(* IEC 61131-3 sources: Industrial-automation-using-LLMs/datasets/Industrial_data/test_harness/test_case (part 2) *)

(* ---- SEQUENCE_8_TestCases (1).st ---- *)
FUNCTION_BLOCK FB_TEST_0
  VAR_OUTPUT
    Finished : BOOL;
    Failed : BOOL;
  END_VAR
  VAR
    TestBlock : SEQUENCE_8;
    TestState : INT;
    Timer : TON;
  END_VAR

  Timer(IN:=TRUE, PT:= T#0s); (* placeholder for later usage *)

  CASE testState OF
    0:
      IF (Timer.Q) THEN
        TestBlock(IN0 := TRUE, IN1 := TRUE, IN2 := TRUE, IN3 := TRUE, IN4 := TRUE, IN5 := TRUE, IN6 := TRUE, IN7 := TRUE, START := FALSE, RST := TRUE, STOP_ON_ERROR := TRUE);
        TestState:=TestState+1;
      END_IF;
      Timer(IN:=TRUE, PT:=T#0s);
    1:
      IF (Timer.Q) THEN
      {printf("0,0: TestBlock.Q0 = FALSE  actual=%lf\n", (double)__GET_VAR(data__->TESTBLOCK.Q0,));}
      {printf("0,0: TestBlock.Q1 = FALSE  actual=%lf\n", (double)__GET_VAR(data__->TESTBLOCK.Q1,));}
      {printf("0,0: TestBlock.Q2 = FALSE  actual=%lf\n", (double)__GET_VAR(data__->TESTBLOCK.Q2,));}
      {printf("0,0: TestBlock.Q3 = FALSE  actual=%lf\n", (double)__GET_VAR(data__->TESTBLOCK.Q3,));}
      {printf("0,0: TestBlock.Q4 = FALSE  actual=%lf\n", (double)__GET_VAR(data__->TESTBLOCK.Q4,));}
      {printf("0,0: TestBlock.Q5 = FALSE  actual=%lf\n", (double)__GET_VAR(data__->TESTBLOCK.Q5,));}
      {printf("0,0: TestBlock.Q6 = FALSE  actual=%lf\n", (double)__GET_VAR(data__->TESTBLOCK.Q6,));}
      {printf("0,0: TestBlock.Q7 = FALSE  actual=%lf\n", (double)__GET_VAR(data__->TESTBLOCK.Q7,));}
      {printf("0,0: TestBlock.QX = FALSE  actual=%lf\n", (double)__GET_VAR(data__->TESTBLOCK.QX,));}
      {printf("0,0: TestBlock.RUN = FALSE  actual=%lf\n", (double)__GET_VAR(data__->TESTBLOCK.RUN,));}
      {printf("0,0: TestBlock._STEP = -1  actual=%lf\n", (double)__GET_VAR(data__->TESTBLOCK._STEP,));}
      {printf("0,0: TestBlock.STATUS = 110  actual=%lf\n", (double)__GET_VAR(data__->TESTBLOCK.STATUS,));}
        IF NOT(TestBlock.Q0 = FALSE AND TestBlock.Q1 = FALSE AND TestBlock.Q2 = FALSE AND TestBlock.Q3 = FALSE AND TestBlock.Q4 = FALSE AND TestBlock.Q5 = FALSE AND TestBlock.Q6 = FALSE AND TestBlock.Q7 = FALSE AND TestBlock.QX = FALSE AND TestBlock.RUN = FALSE AND TestBlock._STEP = -1 AND TestBlock.STATUS = 110) THEN Failed := TRUE; END_IF;
      END_IF;
      Finished:=TRUE;
  END_CASE;
END_FUNCTION_BLOCK

FUNCTION_BLOCK FB_TEST_1
  VAR_OUTPUT
    Finished : BOOL;
    Failed : BOOL;
  END_VAR
  VAR
    TestBlock : SEQUENCE_8;
    TestState : INT;
    Timer : TON;
  END_VAR

  Timer(IN:=TRUE, PT:= T#0s); (* placeholder for later usage *)

  CASE testState OF
    0:
      IF (Timer.Q) THEN
        TestBlock(IN0 := TRUE, IN1 := TRUE, IN2 := TRUE, IN3 := TRUE, IN4 := TRUE, IN5 := TRUE, IN6 := TRUE, IN7 := TRUE, START := TRUE, RST := FALSE, STOP_ON_ERROR := FALSE);
        TestState:=TestState+1;
      END_IF;
      Timer(IN:=TRUE, PT:=T#0s);
    1:
      IF (Timer.Q) THEN
      {printf("1,0: TestBlock.Q0 = TRUE  actual=%lf\n", (double)__GET_VAR(data__->TESTBLOCK.Q0,));}
      {printf("1,0: TestBlock.Q1 = FALSE  actual=%lf\n", (double)__GET_VAR(data__->TESTBLOCK.Q1,));}
      {printf("1,0: TestBlock.Q2 = FALSE  actual=%lf\n", (double)__GET_VAR(data__->TESTBLOCK.Q2,));}
      {printf("1,0: TestBlock.Q3 = FALSE  actual=%lf\n", (double)__GET_VAR(data__->TESTBLOCK.Q3,));}
      {printf("1,0: TestBlock.Q4 = FALSE  actual=%lf\n", (double)__GET_VAR(data__->TESTBLOCK.Q4,));}
      {printf("1,0: TestBlock.Q5 = FALSE  actual=%lf\n", (double)__GET_VAR(data__->TESTBLOCK.Q5,));}
      {printf("1,0: TestBlock.Q6 = FALSE  actual=%lf\n", (double)__GET_VAR(data__->TESTBLOCK.Q6,));}
      {printf("1,0: TestBlock.Q7 = FALSE  actual=%lf\n", (double)__GET_VAR(data__->TESTBLOCK.Q7,));}
      {printf("1,0: TestBlock.QX = TRUE  actual=%lf\n", (double)__GET_VAR(data__->TESTBLOCK.QX,));}
      {printf("1,0: TestBlock.RUN = TRUE  actual=%lf\n", (double)__GET_VAR(data__->TESTBLOCK.RUN,));}
      {printf("1,0: TestBlock._STEP = 0  actual=%lf\n", (double)__GET_VAR(data__->TESTBLOCK._STEP,));}
      {printf("1,0: TestBlock.STATUS = 111  actual=%lf\n", (double)__GET_VAR(data__->TESTBLOCK.STATUS,));}
        IF NOT(TestBlock.Q0 = TRUE AND TestBlock.Q1 = FALSE AND TestBlock.Q2 = FALSE AND TestBlock.Q3 = FALSE AND TestBlock.Q4 = FALSE AND TestBlock.Q5 = FALSE AND TestBlock.Q6 = FALSE AND TestBlock.Q7 = FALSE AND TestBlock.QX = TRUE AND TestBlock.RUN = TRUE AND TestBlock._STEP = 0 AND TestBlock.STATUS = 111) THEN Failed := TRUE; END_IF;
      END_IF;
      Finished:=TRUE;
  END_CASE;
END_FUNCTION_BLOCK

PROGRAM TestRunnerProgram
VAR
  testResult AT %QX0.0 : BOOL := FALSE;
END_VAR
VAR
  totalTests AT %QW0 : INT := 0;
  passedTests AT %QW1 : INT := 0;
END_VAR
VAR
  i: INT := 0;
  testOutcomeArray : ARRAY [0..1] OF BOOL;
  Test_0: FB_TEST_0;
  Test_1: FB_TEST_1;
END_VAR

  IF NOT Test_0.Finished AND NOT Test_0.FAILED THEN totalTests := totalTests + 1; Test_0(); END_IF;
  IF Test_0.Finished THEN testOutcomeArray[0] := TRUE; END_IF;
  IF NOT Test_1.Finished AND NOT Test_1.FAILED THEN totalTests := totalTests + 1; Test_1(); END_IF;
  IF Test_1.Finished THEN testOutcomeArray[1] := TRUE; END_IF;

  passedTests := 0;
  FOR i:=0 TO 1 DO
    IF testOutcomeArray[i]=TRUE THEN passedTests := passedTests+1; END_IF;
  END_FOR;
END_PROGRAM

(* ---- SEQUENCE_8_TestCases.st ---- *)
FUNCTION_BLOCK FB_TEST_0
  VAR_OUTPUT
    Finished : BOOL;
    Failed : BOOL;
  END_VAR
  VAR
    TestBlock : SEQUENCE_8;
    TestState : INT;
    Timer : TON;
  END_VAR

  Timer(IN:=TRUE, PT:= T#0s); (* placeholder for later usage *)

  CASE testState OF
    0:
      IF (Timer.Q) THEN
        TestBlock(IN0 := TRUE, IN1 := TRUE, IN2 := TRUE, IN3 := TRUE, IN4 := TRUE, IN5 := TRUE, IN6 := TRUE, IN7 := TRUE, START := TRUE, RST := FALSE, WAIT0 := T#5s, DELAY0 := T#1s, WAIT1 := T#5s, DELAY1 := T#1s, WAIT2 := T#5s, DELAY2 := T#1s, WAIT3 := T#5s, DELAY3 := T#1s, WAIT4 := T#5s, DELAY4 := T#1s, WAIT5 := T#5s, DELAY5 := T#1s, WAIT6 := T#5s, DELAY6 := T#1s, WAIT7 := T#5s, DELAY7 := T#1s, STOP_ON_ERROR := FALSE);
        TestState:=TestState+1;
      END_IF;
      Timer(IN:=TRUE, PT:=T#0s);
    1:
      IF (Timer.Q) THEN
      {printf("0,0: TestBlock.Q0 = FALSE  actual=%lf\n", (double)__GET_VAR(data__->TESTBLOCK.Q0,));}
      {printf("0,0: TestBlock.Q1 = FALSE  actual=%lf\n", (double)__GET_VAR(data__->TESTBLOCK.Q1,));}
      {printf("0,0: TestBlock.Q2 = FALSE  actual=%lf\n", (double)__GET_VAR(data__->TESTBLOCK.Q2,));}
      {printf("0,0: TestBlock.Q3 = FALSE  actual=%lf\n", (double)__GET_VAR(data__->TESTBLOCK.Q3,));}
      {printf("0,0: TestBlock.Q4 = FALSE  actual=%lf\n", (double)__GET_VAR(data__->TESTBLOCK.Q4,));}
      {printf("0,0: TestBlock.Q5 = FALSE  actual=%lf\n", (double)__GET_VAR(data__->TESTBLOCK.Q5,));}
      {printf("0,0: TestBlock.Q6 = FALSE  actual=%lf\n", (double)__GET_VAR(data__->TESTBLOCK.Q6,));}
      {printf("0,0: TestBlock.Q7 = FALSE  actual=%lf\n", (double)__GET_VAR(data__->TESTBLOCK.Q7,));}
      {printf("0,0: TestBlock.QX = FALSE  actual=%lf\n", (double)__GET_VAR(data__->TESTBLOCK.QX,));}
      {printf("0,0: TestBlock.RUN = FALSE  actual=%lf\n", (double)__GET_VAR(data__->TESTBLOCK.RUN,));}
      {printf("0,0: TestBlock._STEP = -1  actual=%lf\n", (double)__GET_VAR(data__->TESTBLOCK._STEP,));}
      {printf("0,0: TestBlock.STATUS = 110  actual=%lf\n", (double)__GET_VAR(data__->TESTBLOCK.STATUS,));}
        IF NOT(TestBlock.Q0 = FALSE AND TestBlock.Q1 = FALSE AND TestBlock.Q2 = FALSE AND TestBlock.Q3 = FALSE AND TestBlock.Q4 = FALSE AND TestBlock.Q5 = FALSE AND TestBlock.Q6 = FALSE AND TestBlock.Q7 = FALSE AND TestBlock.QX = FALSE AND TestBlock.RUN = FALSE AND TestBlock._STEP = -1 AND TestBlock.STATUS = 110) THEN Failed := TRUE; END_IF;
      END_IF;
      Finished:=TRUE;
  END_CASE;
END_FUNCTION_BLOCK

FUNCTION_BLOCK FB_TEST_1
  VAR_OUTPUT
    Finished : BOOL;
    Failed : BOOL;
  END_VAR
  VAR
    TestBlock : SEQUENCE_8;
    TestState : INT;
    Timer : TON;
  END_VAR

  Timer(IN:=TRUE, PT:= T#0s); (* placeholder for later usage *)

  CASE testState OF
    0:
      IF (Timer.Q) THEN
        TestBlock(IN0 := TRUE, IN1 := TRUE, IN2 := TRUE, IN3 := TRUE, IN4 := TRUE, IN5 := TRUE, IN6 := TRUE, IN7 := TRUE, START := FALSE, RST := TRUE, WAIT0 := T#5s, DELAY0 := T#1s, WAIT1 := T#5s, DELAY1 := T#1s, WAIT2 := T#5s, DELAY2 := T#1s, WAIT3 := T#5s, DELAY3 := T#1s, WAIT4 := T#5s, DELAY4 := T#1s, WAIT5 := T#5s, DELAY5 := T#1s, WAIT6 := T#5s, DELAY6 := T#1s, WAIT7 := T#5s, DELAY7 := T#1s, STOP_ON_ERROR := FALSE);
        TestState:=TestState+1;
      END_IF;
      Timer(IN:=TRUE, PT:=T#0s);
    1:
      IF (Timer.Q) THEN
      {printf("1,0: TestBlock.Q0 = FALSE  actual=%lf\n", (double)__GET_VAR(data__->TESTBLOCK.Q0,));}
      {printf("1,0: TestBlock.Q1 = FALSE  actual=%lf\n", (double)__GET_VAR(data__->TESTBLOCK.Q1,));}
      {printf("1,0: TestBlock.Q2 = FALSE  actual=%lf\n", (double)__GET_VAR(data__->TESTBLOCK.Q2,));}
      {printf("1,0: TestBlock.Q3 = FALSE  actual=%lf\n", (double)__GET_VAR(data__->TESTBLOCK.Q3,));}
      {printf("1,0: TestBlock.Q4 = FALSE  actual=%lf\n", (double)__GET_VAR(data__->TESTBLOCK.Q4,));}
      {printf("1,0: TestBlock.Q5 = FALSE  actual=%lf\n", (double)__GET_VAR(data__->TESTBLOCK.Q5,));}
      {printf("1,0: TestBlock.Q6 = FALSE  actual=%lf\n", (double)__GET_VAR(data__->TESTBLOCK.Q6,));}
      {printf("1,0: TestBlock.Q7 = FALSE  actual=%lf\n", (double)__GET_VAR(data__->TESTBLOCK.Q7,));}
      {printf("1,0: TestBlock.QX = FALSE  actual=%lf\n", (double)__GET_VAR(data__->TESTBLOCK.QX,));}
      {printf("1,0: TestBlock.RUN = FALSE  actual=%lf\n", (double)__GET_VAR(data__->TESTBLOCK.RUN,));}
      {printf("1,0: TestBlock._STEP = -1  actual=%lf\n", (double)__GET_VAR(data__->TESTBLOCK._STEP,));}
      {printf("1,0: TestBlock.STATUS = 110  actual=%lf\n", (double)__GET_VAR(data__->TESTBLOCK.STATUS,));}
        IF NOT(TestBlock.Q0 = FALSE AND TestBlock.Q1 = FALSE AND TestBlock.Q2 = FALSE AND TestBlock.Q3 = FALSE AND TestBlock.Q4 = FALSE AND TestBlock.Q5 = FALSE AND TestBlock.Q6 = FALSE AND TestBlock.Q7 = FALSE AND TestBlock.QX = FALSE AND TestBlock.RUN = FALSE AND TestBlock._STEP = -1 AND TestBlock.STATUS = 110) THEN Failed := TRUE; END_IF;
      END_IF;
      Finished:=TRUE;
  END_CASE;
END_FUNCTION_BLOCK

PROGRAM TestRunnerProgram
VAR
  testResult AT %QX0.0 : BOOL := FALSE;
END_VAR
VAR
  totalTests AT %QW0 : INT := 0;
  passedTests AT %QW1 : INT := 0;
END_VAR
VAR
  i: INT := 0;
  testOutcomeArray : ARRAY [0..1] OF BOOL;
  Test_0: FB_TEST_0;
  Test_1: FB_TEST_1;
END_VAR

  IF NOT Test_0.Finished AND NOT Test_0.FAILED THEN totalTests := totalTests + 1; Test_0(); END_IF;
  IF Test_0.Finished THEN testOutcomeArray[0] := TRUE; END_IF;
  IF NOT Test_1.Finished AND NOT Test_1.FAILED THEN totalTests := totalTests + 1; Test_1(); END_IF;
  IF Test_1.Finished THEN testOutcomeArray[1] := TRUE; END_IF;

  passedTests := 0;
  FOR i:=0 TO 1 DO
    IF testOutcomeArray[i]=TRUE THEN passedTests := passedTests+1; END_IF;
  END_FOR;
END_PROGRAM

(* ---- TOOL_CHANGER_TestCases (1).st ---- *)
FUNCTION_BLOCK FB_TEST_0
  VAR_OUTPUT
    Finished : BOOL;
    Failed : BOOL;
  END_VAR
  VAR
    TestBlock : TOOL_CHANGER;
    TestState : INT;
    Timer : TON;
  END_VAR

  Timer(IN:=TRUE, PT:= T#0s); (* placeholder for later usage *)

  CASE testState OF
    0:
      IF (Timer.Q) THEN
        TestBlock(ToolChangeRequired := TRUE, ToolCarouselPosition := 1, DesiredToolNumber := 3);
        TestState:=TestState+1;
      END_IF;
      Timer(IN:=TRUE, PT:=T#0s);
    1:
      IF (Timer.Q) THEN
      {printf("0,0: TestBlock.RotateCarousel = TRUE  actual=%lf\n", (double)__GET_VAR(data__->TESTBLOCK.ROTATECAROUSEL,));}
      {printf("0,0: TestBlock.LockTool = FALSE  actual=%lf\n", (double)__GET_VAR(data__->TESTBLOCK.LOCKTOOL,));}
        IF NOT (TestBlock.RotateCarousel = TRUE AND TestBlock.LockTool = FALSE) THEN Failed := TRUE; END_IF;
        TestBlock(ToolChangeRequired := TRUE, ToolCarouselPosition := 3, DesiredToolNumber := 3);
        TestState:=TestState+1;
      END_IF;
      Timer(IN:=TRUE, PT:=T#0s);
    2:
      IF (Timer.Q) THEN
      {printf("0,1: TestBlock.RotateCarousel = FALSE  actual=%lf\n", (double)__GET_VAR(data__->TESTBLOCK.ROTATECAROUSEL,));}
      {printf("0,1: TestBlock.LockTool = TRUE  actual=%lf\n", (double)__GET_VAR(data__->TESTBLOCK.LOCKTOOL,));}
        IF NOT (TestBlock.RotateCarousel = FALSE AND TestBlock.LockTool = TRUE) THEN Failed := TRUE; END_IF;
        TestBlock(ToolChangeRequired := TRUE, ToolCarouselPosition := 3, DesiredToolNumber := 3);
        TestState:=TestState+1;
      END_IF;
      Timer(IN:=TRUE, PT:=T#0s);
    3:
      IF (Timer.Q) THEN
      {printf("0,2: TestBlock.RotateCarousel = FALSE  actual=%lf\n", (double)__GET_VAR(data__->TESTBLOCK.ROTATECAROUSEL,));}
      {printf("0,2: TestBlock.LockTool = FALSE  actual=%lf\n", (double)__GET_VAR(data__->TESTBLOCK.LOCKTOOL,));}
        IF NOT(TestBlock.RotateCarousel = FALSE AND TestBlock.LockTool = FALSE) THEN Failed := TRUE; END_IF;
      END_IF;
      Finished:=TRUE;
  END_CASE;
END_FUNCTION_BLOCK

FUNCTION_BLOCK FB_TEST_1
  VAR_OUTPUT
    Finished : BOOL;
    Failed : BOOL;
  END_VAR
  VAR
    TestBlock : TOOL_CHANGER;
    TestState : INT;
    Timer : TON;
  END_VAR

  Timer(IN:=TRUE, PT:= T#0s); (* placeholder for later usage *)

  CASE testState OF
    0:
      IF (Timer.Q) THEN
        TestBlock(ToolChangeRequired := TRUE, ToolCarouselPosition := 5, DesiredToolNumber := 5);
        TestState:=TestState+1;
      END_IF;
      Timer(IN:=TRUE, PT:=T#0s);
    1:
      IF (Timer.Q) THEN
      {printf("1,0: TestBlock.RotateCarousel = FALSE  actual=%lf\n", (double)__GET_VAR(data__->TESTBLOCK.ROTATECAROUSEL,));}
      {printf("1,0: TestBlock.LockTool = TRUE  actual=%lf\n", (double)__GET_VAR(data__->TESTBLOCK.LOCKTOOL,));}
        IF NOT (TestBlock.RotateCarousel = FALSE AND TestBlock.LockTool = TRUE) THEN Failed := TRUE; END_IF;
        TestBlock(ToolChangeRequired := TRUE, ToolCarouselPosition := 1, DesiredToolNumber := 1);
        TestState:=TestState+1;
      END_IF;
      Timer(IN:=TRUE, PT:=T#0s);
    2:
      IF (Timer.Q) THEN
      {printf("1,1: TestBlock.RotateCarousel = FALSE  actual=%lf\n", (double)__GET_VAR(data__->TESTBLOCK.ROTATECAROUSEL,));}
      {printf("1,1: TestBlock.LockTool = TRUE  actual=%lf\n", (double)__GET_VAR(data__->TESTBLOCK.LOCKTOOL,));}
        IF NOT (TestBlock.RotateCarousel = FALSE AND TestBlock.LockTool = TRUE) THEN Failed := TRUE; END_IF;
        TestBlock(ToolChangeRequired := TRUE, ToolCarouselPosition := 1, DesiredToolNumber := 1);
        TestState:=TestState+1;
      END_IF;
      Timer(IN:=TRUE, PT:=T#0s);
    3:
      IF (Timer.Q) THEN
      {printf("1,2: TestBlock.RotateCarousel = FALSE  actual=%lf\n", (double)__GET_VAR(data__->TESTBLOCK.ROTATECAROUSEL,));}
      {printf("1,2: TestBlock.LockTool = FALSE  actual=%lf\n", (double)__GET_VAR(data__->TESTBLOCK.LOCKTOOL,));}
        IF NOT(TestBlock.RotateCarousel = FALSE AND TestBlock.LockTool = FALSE) THEN Failed := TRUE; END_IF;
      END_IF;
      Finished:=TRUE;
  END_CASE;
END_FUNCTION_BLOCK

FUNCTION_BLOCK FB_TEST_2
  VAR_OUTPUT
    Finished : BOOL;
    Failed : BOOL;
  END_VAR
  VAR
    TestBlock : TOOL_CHANGER;
    TestState : INT;
    Timer : TON;
  END_VAR

  Timer(IN:=TRUE, PT:= T#0s); (* placeholder for later usage *)

  CASE testState OF
    0:
      IF (Timer.Q) THEN
        TestBlock(ToolChangeRequired := FALSE, ToolCarouselPosition := 2, DesiredToolNumber := 2);
        TestState:=TestState+1;
      END_IF;
      Timer(IN:=TRUE, PT:=T#0s);
    1:
      IF (Timer.Q) THEN
      {printf("2,0: TestBlock.RotateCarousel = FALSE  actual=%lf\n", (double)__GET_VAR(data__->TESTBLOCK.ROTATECAROUSEL,));}
      {printf("2,0: TestBlock.LockTool = FALSE  actual=%lf\n", (double)__GET_VAR(data__->TESTBLOCK.LOCKTOOL,));}
        IF NOT (TestBlock.RotateCarousel = FALSE AND TestBlock.LockTool = FALSE) THEN Failed := TRUE; END_IF;
        TestBlock(ToolChangeRequired := FALSE, ToolCarouselPosition := 2, DesiredToolNumber := 3);
        TestState:=TestState+1;
      END_IF;
      Timer(IN:=TRUE, PT:=T#0s);
    2:
      IF (Timer.Q) THEN
      {printf("2,1: TestBlock.RotateCarousel = FALSE  actual=%lf\n", (double)__GET_VAR(data__->TESTBLOCK.ROTATECAROUSEL,));}
      {printf("2,1: TestBlock.LockTool = FALSE  actual=%lf\n", (double)__GET_VAR(data__->TESTBLOCK.LOCKTOOL,));}
        IF NOT (TestBlock.RotateCarousel = FALSE AND TestBlock.LockTool = FALSE) THEN Failed := TRUE; END_IF;
        TestBlock(ToolChangeRequired := FALSE, ToolCarouselPosition := 3, DesiredToolNumber := 3);
        TestState:=TestState+1;
      END_IF;
      Timer(IN:=TRUE, PT:=T#0s);
    3:
      IF (Timer.Q) THEN
      {printf("2,2: TestBlock.RotateCarousel = FALSE  actual=%lf\n", (double)__GET_VAR(data__->TESTBLOCK.ROTATECAROUSEL,));}
      {printf("2,2: TestBlock.LockTool = FALSE  actual=%lf\n", (double)__GET_VAR(data__->TESTBLOCK.LOCKTOOL,));}
        IF NOT(TestBlock.RotateCarousel = FALSE AND TestBlock.LockTool = FALSE) THEN Failed := TRUE; END_IF;
      END_IF;
      Finished:=TRUE;
  END_CASE;
END_FUNCTION_BLOCK

PROGRAM TestRunnerProgram
VAR
  testResult AT %QX0.0 : BOOL := FALSE;
END_VAR
VAR
  totalTests AT %QW0 : INT := 0;
  passedTests AT %QW1 : INT := 0;
END_VAR
VAR
  i: INT := 0;
  testOutcomeArray : ARRAY [0..2] OF BOOL;
  Test_0: FB_TEST_0;
  Test_1: FB_TEST_1;
  Test_2: FB_TEST_2;
END_VAR

  IF NOT Test_0.Finished AND NOT Test_0.FAILED THEN totalTests := totalTests + 1; Test_0(); END_IF;
  IF Test_0.Finished THEN testOutcomeArray[0] := TRUE; END_IF;
  IF NOT Test_1.Finished AND NOT Test_1.FAILED THEN totalTests := totalTests + 1; Test_1(); END_IF;
  IF Test_1.Finished THEN testOutcomeArray[1] := TRUE; END_IF;
  IF NOT Test_2.Finished AND NOT Test_2.FAILED THEN totalTests := totalTests + 1; Test_2(); END_IF;
  IF Test_2.Finished THEN testOutcomeArray[2] := TRUE; END_IF;

  passedTests := 0;
  FOR i:=0 TO 2 DO
    IF testOutcomeArray[i]=TRUE THEN passedTests := passedTests+1; END_IF;
  END_FOR;
END_PROGRAM

(* ---- TOOL_CHANGER_TestCases.st ---- *)
FUNCTION_BLOCK FB_TEST_0
  VAR_OUTPUT
    Finished : BOOL;
    Failed : BOOL;
  END_VAR
  VAR
    TestBlock : TOOL_CHANGER;
    TestState : INT;
    Timer : TON;
  END_VAR

  Timer(IN:=TRUE, PT:= T#0s); (* placeholder for later usage *)

  CASE testState OF
    0:
      IF (Timer.Q) THEN
        TestBlock(ToolChangeRequired := TRUE, ToolCarouselPosition := 1, DesiredToolNumber := 2);
        TestState:=TestState+1;
      END_IF;
      Timer(IN:=TRUE, PT:=T#0s);
    1:
      IF (Timer.Q) THEN
      {printf("0,0: TestBlock.RotateCarousel = TRUE  actual=%lf\n", (double)__GET_VAR(data__->TESTBLOCK.ROTATECAROUSEL,));}
      {printf("0,0: TestBlock.LockTool = FALSE  actual=%lf\n", (double)__GET_VAR(data__->TESTBLOCK.LOCKTOOL,));}
        IF NOT(TestBlock.RotateCarousel = TRUE AND TestBlock.LockTool = FALSE) THEN Failed := TRUE; END_IF;
      END_IF;
      Finished:=TRUE;
  END_CASE;
END_FUNCTION_BLOCK

FUNCTION_BLOCK FB_TEST_1
  VAR_OUTPUT
    Finished : BOOL;
    Failed : BOOL;
  END_VAR
  VAR
    TestBlock : TOOL_CHANGER;
    TestState : INT;
    Timer : TON;
  END_VAR

  Timer(IN:=TRUE, PT:= T#0s); (* placeholder for later usage *)

  CASE testState OF
    0:
      IF (Timer.Q) THEN
        TestBlock(ToolChangeRequired := TRUE, ToolCarouselPosition := 2, DesiredToolNumber := 2);
        TestState:=TestState+1;
      END_IF;
      Timer(IN:=TRUE, PT:=T#0s);
    1:
      IF (Timer.Q) THEN
      {printf("1,0: TestBlock.RotateCarousel = FALSE  actual=%lf\n", (double)__GET_VAR(data__->TESTBLOCK.ROTATECAROUSEL,));}
      {printf("1,0: TestBlock.LockTool = TRUE  actual=%lf\n", (double)__GET_VAR(data__->TESTBLOCK.LOCKTOOL,));}
        IF NOT(TestBlock.RotateCarousel = FALSE AND TestBlock.LockTool = TRUE) THEN Failed := TRUE; END_IF;
      END_IF;
      Finished:=TRUE;
  END_CASE;
END_FUNCTION_BLOCK

FUNCTION_BLOCK FB_TEST_2
  VAR_OUTPUT
    Finished : BOOL;
    Failed : BOOL;
  END_VAR
  VAR
    TestBlock : TOOL_CHANGER;
    TestState : INT;
    Timer : TON;
  END_VAR

  Timer(IN:=TRUE, PT:= T#0s); (* placeholder for later usage *)

  CASE testState OF
    0:
      IF (Timer.Q) THEN
        TestBlock(ToolChangeRequired := TRUE, ToolCarouselPosition := 2, DesiredToolNumber := 1);
        TestState:=TestState+1;
      END_IF;
      Timer(IN:=TRUE, PT:=T#0s);
    1:
      IF (Timer.Q) THEN
      {printf("2,0: TestBlock.RotateCarousel = TRUE  actual=%lf\n", (double)__GET_VAR(data__->TESTBLOCK.ROTATECAROUSEL,));}
      {printf("2,0: TestBlock.LockTool = FALSE  actual=%lf\n", (double)__GET_VAR(data__->TESTBLOCK.LOCKTOOL,));}
        IF NOT(TestBlock.RotateCarousel = TRUE AND TestBlock.LockTool = FALSE) THEN Failed := TRUE; END_IF;
      END_IF;
      Finished:=TRUE;
  END_CASE;
END_FUNCTION_BLOCK

FUNCTION_BLOCK FB_TEST_3
  VAR_OUTPUT
    Finished : BOOL;
    Failed : BOOL;
  END_VAR
  VAR
    TestBlock : TOOL_CHANGER;
    TestState : INT;
    Timer : TON;
  END_VAR

  Timer(IN:=TRUE, PT:= T#0s); (* placeholder for later usage *)

  CASE testState OF
    0:
      IF (Timer.Q) THEN
        TestBlock(ToolChangeRequired := FALSE, ToolCarouselPosition := 1, DesiredToolNumber := 1);
        TestState:=TestState+1;
      END_IF;
      Timer(IN:=TRUE, PT:=T#0s);
    1:
      IF (Timer.Q) THEN
      {printf("3,0: TestBlock.RotateCarousel = FALSE  actual=%lf\n", (double)__GET_VAR(data__->TESTBLOCK.ROTATECAROUSEL,));}
      {printf("3,0: TestBlock.LockTool = FALSE  actual=%lf\n", (double)__GET_VAR(data__->TESTBLOCK.LOCKTOOL,));}
        IF NOT(TestBlock.RotateCarousel = FALSE AND TestBlock.LockTool = FALSE) THEN Failed := TRUE; END_IF;
      END_IF;
      Finished:=TRUE;
  END_CASE;
END_FUNCTION_BLOCK

FUNCTION_BLOCK FB_TEST_4
  VAR_OUTPUT
    Finished : BOOL;
    Failed : BOOL;
  END_VAR
  VAR
    TestBlock : TOOL_CHANGER;
    TestState : INT;
    Timer : TON;
  END_VAR

  Timer(IN:=TRUE, PT:= T#0s); (* placeholder for later usage *)

  CASE testState OF
    0:
      IF (Timer.Q) THEN
        TestBlock(ToolChangeRequired := FALSE, ToolCarouselPosition := 1, DesiredToolNumber := 2);
        TestState:=TestState+1;
      END_IF;
      Timer(IN:=TRUE, PT:=T#0s);
    1:
      IF (Timer.Q) THEN
      {printf("4,0: TestBlock.RotateCarousel = FALSE  actual=%lf\n", (double)__GET_VAR(data__->TESTBLOCK.ROTATECAROUSEL,));}
      {printf("4,0: TestBlock.LockTool = FALSE  actual=%lf\n", (double)__GET_VAR(data__->TESTBLOCK.LOCKTOOL,));}
        IF NOT(TestBlock.RotateCarousel = FALSE AND TestBlock.LockTool = FALSE) THEN Failed := TRUE; END_IF;
      END_IF;
      Finished:=TRUE;
  END_CASE;
END_FUNCTION_BLOCK

PROGRAM TestRunnerProgram
VAR
  testResult AT %QX0.0 : BOOL := FALSE;
END_VAR
VAR
  totalTests AT %QW0 : INT := 0;
  passedTests AT %QW1 : INT := 0;
END_VAR
VAR
  i: INT := 0;
  testOutcomeArray : ARRAY [0..4] OF BOOL;
  Test_0: FB_TEST_0;
  Test_1: FB_TEST_1;
  Test_2: FB_TEST_2;
  Test_3: FB_TEST_3;
  Test_4: FB_TEST_4;
END_VAR

  IF NOT Test_0.Finished AND NOT Test_0.FAILED THEN totalTests := totalTests + 1; Test_0(); END_IF;
  IF Test_0.Finished THEN testOutcomeArray[0] := TRUE; END_IF;
  IF NOT Test_1.Finished AND NOT Test_1.FAILED THEN totalTests := totalTests + 1; Test_1(); END_IF;
  IF Test_1.Finished THEN testOutcomeArray[1] := TRUE; END_IF;
  IF NOT Test_2.Finished AND NOT Test_2.FAILED THEN totalTests := totalTests + 1; Test_2(); END_IF;
  IF Test_2.Finished THEN testOutcomeArray[2] := TRUE; END_IF;
  IF NOT Test_3.Finished AND NOT Test_3.FAILED THEN totalTests := totalTests + 1; Test_3(); END_IF;
  IF Test_3.Finished THEN testOutcomeArray[3] := TRUE; END_IF;
  IF NOT Test_4.Finished AND NOT Test_4.FAILED THEN totalTests := totalTests + 1; Test_4(); END_IF;
  IF Test_4.Finished THEN testOutcomeArray[4] := TRUE; END_IF;

  passedTests := 0;
  FOR i:=0 TO 4 DO
    IF testOutcomeArray[i]=TRUE THEN passedTests := passedTests+1; END_IF;
  END_FOR;
END_PROGRAM

(* ---- TRAFFIC_CTRL_TestCases (1).st ---- *)
FUNCTION_BLOCK FB_TEST_0
  VAR_OUTPUT
    Finished : BOOL;
    Failed : BOOL;
  END_VAR
  VAR
    TestBlock : TRAFFIC_CTRL;
    TestState : INT;
    Timer : TON;
  END_VAR

  Timer(IN:=TRUE, PT:= T#0s); (* placeholder for later usage *)

  CASE testState OF
    0:
      IF (Timer.Q) THEN
        TestBlock(PedestrianButton1 := FALSE, PedestrianButton2 := FALSE);
        TestState:=TestState+1;
      END_IF;
      Timer(IN:=TRUE, PT:=T#0s);
    1:
      IF (Timer.Q) THEN
      {printf("0,0: TestBlock.NorthSouthRed = FALSE  actual=%lf\n", (double)__GET_VAR(data__->TESTBLOCK.NORTHSOUTHRED,));}
      {printf("0,0: TestBlock.NorthSouthYellow = FALSE  actual=%lf\n", (double)__GET_VAR(data__->TESTBLOCK.NORTHSOUTHYELLOW,));}
      {printf("0,0: TestBlock.NorthSouthGreen = TRUE  actual=%lf\n", (double)__GET_VAR(data__->TESTBLOCK.NORTHSOUTHGREEN,));}
      {printf("0,0: TestBlock.EastWestRed = TRUE  actual=%lf\n", (double)__GET_VAR(data__->TESTBLOCK.EASTWESTRED,));}
      {printf("0,0: TestBlock.EastWestYellow = FALSE  actual=%lf\n", (double)__GET_VAR(data__->TESTBLOCK.EASTWESTYELLOW,));}
      {printf("0,0: TestBlock.EastWestGreen = FALSE  actual=%lf\n", (double)__GET_VAR(data__->TESTBLOCK.EASTWESTGREEN,));}
      {printf("0,0: TestBlock.PedestrianLight1 = FALSE  actual=%lf\n", (double)__GET_VAR(data__->TESTBLOCK.PEDESTRIANLIGHT1,));}
      {printf("0,0: TestBlock.PedestrianLight2 = FALSE  actual=%lf\n", (double)__GET_VAR(data__->TESTBLOCK.PEDESTRIANLIGHT2,));}
        IF NOT (TestBlock.NorthSouthRed = FALSE AND TestBlock.NorthSouthYellow = FALSE AND TestBlock.NorthSouthGreen = TRUE AND TestBlock.EastWestRed = TRUE AND TestBlock.EastWestYellow = FALSE AND TestBlock.EastWestGreen = FALSE AND TestBlock.PedestrianLight1 = FALSE AND TestBlock.PedestrianLight2 = FALSE) THEN Failed := TRUE; END_IF;
        TestBlock(PedestrianButton1 := TRUE, PedestrianButton2 := FALSE);
        TestState:=TestState+1;
      END_IF;
      Timer(IN:=TRUE, PT:=T#0s);
    2:
      IF (Timer.Q) THEN
      {printf("0,1: TestBlock.NorthSouthRed = FALSE  actual=%lf\n", (double)__GET_VAR(data__->TESTBLOCK.NORTHSOUTHRED,));}
      {printf("0,1: TestBlock.NorthSouthYellow = TRUE  actual=%lf\n", (double)__GET_VAR(data__->TESTBLOCK.NORTHSOUTHYELLOW,));}
      {printf("0,1: TestBlock.NorthSouthGreen = FALSE  actual=%lf\n", (double)__GET_VAR(data__->TESTBLOCK.NORTHSOUTHGREEN,));}
      {printf("0,1: TestBlock.EastWestRed = TRUE  actual=%lf\n", (double)__GET_VAR(data__->TESTBLOCK.EASTWESTRED,));}
      {printf("0,1: TestBlock.EastWestYellow = FALSE  actual=%lf\n", (double)__GET_VAR(data__->TESTBLOCK.EASTWESTYELLOW,));}
      {printf("0,1: TestBlock.EastWestGreen = FALSE  actual=%lf\n", (double)__GET_VAR(data__->TESTBLOCK.EASTWESTGREEN,));}
      {printf("0,1: TestBlock.PedestrianLight1 = FALSE  actual=%lf\n", (double)__GET_VAR(data__->TESTBLOCK.PEDESTRIANLIGHT1,));}
      {printf("0,1: TestBlock.PedestrianLight2 = FALSE  actual=%lf\n", (double)__GET_VAR(data__->TESTBLOCK.PEDESTRIANLIGHT2,));}
        IF NOT(TestBlock.NorthSouthRed = FALSE AND TestBlock.NorthSouthYellow = TRUE AND TestBlock.NorthSouthGreen = FALSE AND TestBlock.EastWestRed = TRUE AND TestBlock.EastWestYellow = FALSE AND TestBlock.EastWestGreen = FALSE AND TestBlock.PedestrianLight1 = FALSE AND TestBlock.PedestrianLight2 = FALSE) THEN Failed := TRUE; END_IF;
      END_IF;
      Finished:=TRUE;
  END_CASE;
END_FUNCTION_BLOCK

FUNCTION_BLOCK FB_TEST_1
  VAR_OUTPUT
    Finished : BOOL;
    Failed : BOOL;
  END_VAR
  VAR
    TestBlock : TRAFFIC_CTRL;
    TestState : INT;
    Timer : TON;
  END_VAR

  Timer(IN:=TRUE, PT:= T#0s); (* placeholder for later usage *)

  CASE testState OF
    0:
      IF (Timer.Q) THEN
        TestBlock(PedestrianButton1 := FALSE, PedestrianButton2 := TRUE);
        TestState:=TestState+1;
      END_IF;
      Timer(IN:=TRUE, PT:=T#0s);
    1:
      IF (Timer.Q) THEN
      {printf("1,0: TestBlock.NorthSouthRed = TRUE  actual=%lf\n", (double)__GET_VAR(data__->TESTBLOCK.NORTHSOUTHRED,));}
      {printf("1,0: TestBlock.NorthSouthYellow = FALSE  actual=%lf\n", (double)__GET_VAR(data__->TESTBLOCK.NORTHSOUTHYELLOW,));}
      {printf("1,0: TestBlock.NorthSouthGreen = FALSE  actual=%lf\n", (double)__GET_VAR(data__->TESTBLOCK.NORTHSOUTHGREEN,));}
      {printf("1,0: TestBlock.EastWestRed = FALSE  actual=%lf\n", (double)__GET_VAR(data__->TESTBLOCK.EASTWESTRED,));}
      {printf("1,0: TestBlock.EastWestYellow = FALSE  actual=%lf\n", (double)__GET_VAR(data__->TESTBLOCK.EASTWESTYELLOW,));}
      {printf("1,0: TestBlock.EastWestGreen = TRUE  actual=%lf\n", (double)__GET_VAR(data__->TESTBLOCK.EASTWESTGREEN,));}
      {printf("1,0: TestBlock.PedestrianLight1 = FALSE  actual=%lf\n", (double)__GET_VAR(data__->TESTBLOCK.PEDESTRIANLIGHT1,));}
      {printf("1,0: TestBlock.PedestrianLight2 = TRUE  actual=%lf\n", (double)__GET_VAR(data__->TESTBLOCK.PEDESTRIANLIGHT2,));}
        IF NOT (TestBlock.NorthSouthRed = TRUE AND TestBlock.NorthSouthYellow = FALSE AND TestBlock.NorthSouthGreen = FALSE AND TestBlock.EastWestRed = FALSE AND TestBlock.EastWestYellow = FALSE AND TestBlock.EastWestGreen = TRUE AND TestBlock.PedestrianLight1 = FALSE AND TestBlock.PedestrianLight2 = TRUE) THEN Failed := TRUE; END_IF;
        TestBlock(PedestrianButton1 := FALSE, PedestrianButton2 := FALSE);
        TestState:=TestState+1;
      END_IF;
      Timer(IN:=TRUE, PT:=T#0s);
    2:
      IF (Timer.Q) THEN
      {printf("1,1: TestBlock.NorthSouthRed = TRUE  actual=%lf\n", (double)__GET_VAR(data__->TESTBLOCK.NORTHSOUTHRED,));}
      {printf("1,1: TestBlock.NorthSouthYellow = FALSE  actual=%lf\n", (double)__GET_VAR(data__->TESTBLOCK.NORTHSOUTHYELLOW,));}
      {printf("1,1: TestBlock.NorthSouthGreen = FALSE  actual=%lf\n", (double)__GET_VAR(data__->TESTBLOCK.NORTHSOUTHGREEN,));}
      {printf("1,1: TestBlock.EastWestRed = FALSE  actual=%lf\n", (double)__GET_VAR(data__->TESTBLOCK.EASTWESTRED,));}
      {printf("1,1: TestBlock.EastWestYellow = TRUE  actual=%lf\n", (double)__GET_VAR(data__->TESTBLOCK.EASTWESTYELLOW,));}
      {printf("1,1: TestBlock.EastWestGreen = FALSE  actual=%lf\n", (double)__GET_VAR(data__->TESTBLOCK.EASTWESTGREEN,));}
      {printf("1,1: TestBlock.PedestrianLight1 = FALSE  actual=%lf\n", (double)__GET_VAR(data__->TESTBLOCK.PEDESTRIANLIGHT1,));}
      {printf("1,1: TestBlock.PedestrianLight2 = FALSE  actual=%lf\n", (double)__GET_VAR(data__->TESTBLOCK.PEDESTRIANLIGHT2,));}
        IF NOT(TestBlock.NorthSouthRed = TRUE AND TestBlock.NorthSouthYellow = FALSE AND TestBlock.NorthSouthGreen = FALSE AND TestBlock.EastWestRed = FALSE AND TestBlock.EastWestYellow = TRUE AND TestBlock.EastWestGreen = FALSE AND TestBlock.PedestrianLight1 = FALSE AND TestBlock.PedestrianLight2 = FALSE) THEN Failed := TRUE; END_IF;
      END_IF;
      Finished:=TRUE;
  END_CASE;
END_FUNCTION_BLOCK

PROGRAM TestRunnerProgram
VAR
  testResult AT %QX0.0 : BOOL := FALSE;
END_VAR
VAR
  totalTests AT %QW0 : INT := 0;
  passedTests AT %QW1 : INT := 0;
END_VAR
VAR
  i: INT := 0;
  testOutcomeArray : ARRAY [0..1] OF BOOL;
  Test_0: FB_TEST_0;
  Test_1: FB_TEST_1;
END_VAR

  IF NOT Test_0.Finished AND NOT Test_0.FAILED THEN totalTests := totalTests + 1; Test_0(); END_IF;
  IF Test_0.Finished THEN testOutcomeArray[0] := TRUE; END_IF;
  IF NOT Test_1.Finished AND NOT Test_1.FAILED THEN totalTests := totalTests + 1; Test_1(); END_IF;
  IF Test_1.Finished THEN testOutcomeArray[1] := TRUE; END_IF;

  passedTests := 0;
  FOR i:=0 TO 1 DO
    IF testOutcomeArray[i]=TRUE THEN passedTests := passedTests+1; END_IF;
  END_FOR;
END_PROGRAM

(* ---- TRAFFIC_CTRL_TestCases.st ---- *)
FUNCTION_BLOCK FB_TEST_0
  VAR_OUTPUT
    Finished : BOOL;
    Failed : BOOL;
  END_VAR
  VAR
    TestBlock : TRAFFIC_CTRL;
    TestState : INT;
    Timer : TON;
  END_VAR

  Timer(IN:=TRUE, PT:= T#0s); (* placeholder for later usage *)

  CASE testState OF
    0:
      IF (Timer.Q) THEN
        TestBlock(PedestrianButton1 := FALSE, PedestrianButton2 := FALSE);
        TestState:=TestState+1;
      END_IF;
      Timer(IN:=TRUE, PT:=T#0s);
    1:
      IF (Timer.Q) THEN
      {printf("0,0: TestBlock.NorthSouthRed = FALSE  actual=%lf\n", (double)__GET_VAR(data__->TESTBLOCK.NORTHSOUTHRED,));}
      {printf("0,0: TestBlock.NorthSouthYellow = FALSE  actual=%lf\n", (double)__GET_VAR(data__->TESTBLOCK.NORTHSOUTHYELLOW,));}
      {printf("0,0: TestBlock.NorthSouthGreen = TRUE  actual=%lf\n", (double)__GET_VAR(data__->TESTBLOCK.NORTHSOUTHGREEN,));}
      {printf("0,0: TestBlock.EastWestRed = TRUE  actual=%lf\n", (double)__GET_VAR(data__->TESTBLOCK.EASTWESTRED,));}
      {printf("0,0: TestBlock.EastWestYellow = FALSE  actual=%lf\n", (double)__GET_VAR(data__->TESTBLOCK.EASTWESTYELLOW,));}
      {printf("0,0: TestBlock.EastWestGreen = FALSE  actual=%lf\n", (double)__GET_VAR(data__->TESTBLOCK.EASTWESTGREEN,));}
      {printf("0,0: TestBlock.PedestrianLight1 = FALSE  actual=%lf\n", (double)__GET_VAR(data__->TESTBLOCK.PEDESTRIANLIGHT1,));}
      {printf("0,0: TestBlock.PedestrianLight2 = FALSE  actual=%lf\n", (double)__GET_VAR(data__->TESTBLOCK.PEDESTRIANLIGHT2,));}
        IF NOT(TestBlock.NorthSouthRed = FALSE AND TestBlock.NorthSouthYellow = FALSE AND TestBlock.NorthSouthGreen = TRUE AND TestBlock.EastWestRed = TRUE AND TestBlock.EastWestYellow = FALSE AND TestBlock.EastWestGreen = FALSE AND TestBlock.PedestrianLight1 = FALSE AND TestBlock.PedestrianLight2 = FALSE) THEN Failed := TRUE; END_IF;
      END_IF;
      Finished:=TRUE;
  END_CASE;
END_FUNCTION_BLOCK

FUNCTION_BLOCK FB_TEST_1
  VAR_OUTPUT
    Finished : BOOL;
    Failed : BOOL;
  END_VAR
  VAR
    TestBlock : TRAFFIC_CTRL;
    TestState : INT;
    Timer : TON;
  END_VAR

  Timer(IN:=TRUE, PT:= T#0s); (* placeholder for later usage *)

  CASE testState OF
    0:
      IF (Timer.Q) THEN
        TestBlock(PedestrianButton1 := TRUE, PedestrianButton2 := FALSE);
        TestState:=TestState+1;
      END_IF;
      Timer(IN:=TRUE, PT:=T#0s);
    1:
      IF (Timer.Q) THEN
      {printf("1,0: TestBlock.NorthSouthRed = FALSE  actual=%lf\n", (double)__GET_VAR(data__->TESTBLOCK.NORTHSOUTHRED,));}
      {printf("1,0: TestBlock.NorthSouthYellow = TRUE  actual=%lf\n", (double)__GET_VAR(data__->TESTBLOCK.NORTHSOUTHYELLOW,));}
      {printf("1,0: TestBlock.NorthSouthGreen = FALSE  actual=%lf\n", (double)__GET_VAR(data__->TESTBLOCK.NORTHSOUTHGREEN,));}
      {printf("1,0: TestBlock.EastWestRed = TRUE  actual=%lf\n", (double)__GET_VAR(data__->TESTBLOCK.EASTWESTRED,));}
      {printf("1,0: TestBlock.EastWestYellow = FALSE  actual=%lf\n", (double)__GET_VAR(data__->TESTBLOCK.EASTWESTYELLOW,));}
      {printf("1,0: TestBlock.EastWestGreen = FALSE  actual=%lf\n", (double)__GET_VAR(data__->TESTBLOCK.EASTWESTGREEN,));}
      {printf("1,0: TestBlock.PedestrianLight1 = FALSE  actual=%lf\n", (double)__GET_VAR(data__->TESTBLOCK.PEDESTRIANLIGHT1,));}
      {printf("1,0: TestBlock.PedestrianLight2 = FALSE  actual=%lf\n", (double)__GET_VAR(data__->TESTBLOCK.PEDESTRIANLIGHT2,));}
        IF NOT(TestBlock.NorthSouthRed = FALSE AND TestBlock.NorthSouthYellow = TRUE AND TestBlock.NorthSouthGreen = FALSE AND TestBlock.EastWestRed = TRUE AND TestBlock.EastWestYellow = FALSE AND TestBlock.EastWestGreen = FALSE AND TestBlock.PedestrianLight1 = FALSE AND TestBlock.PedestrianLight2 = FALSE) THEN Failed := TRUE; END_IF;
      END_IF;
      Finished:=TRUE;
  END_CASE;
END_FUNCTION_BLOCK

FUNCTION_BLOCK FB_TEST_2
  VAR_OUTPUT
    Finished : BOOL;
    Failed : BOOL;
  END_VAR
  VAR
    TestBlock : TRAFFIC_CTRL;
    TestState : INT;
    Timer : TON;
  END_VAR

  Timer(IN:=TRUE, PT:= T#0s); (* placeholder for later usage *)

  CASE testState OF
    0:
      IF (Timer.Q) THEN
        TestBlock(PedestrianButton1 := FALSE, PedestrianButton2 := TRUE);
        TestState:=TestState+1;
      END_IF;
      Timer(IN:=TRUE, PT:=T#0s);
    1:
      IF (Timer.Q) THEN
      {printf("2,0: TestBlock.NorthSouthRed = TRUE  actual=%lf\n", (double)__GET_VAR(data__->TESTBLOCK.NORTHSOUTHRED,));}
      {printf("2,0: TestBlock.NorthSouthYellow = FALSE  actual=%lf\n", (double)__GET_VAR(data__->TESTBLOCK.NORTHSOUTHYELLOW,));}
      {printf("2,0: TestBlock.NorthSouthGreen = FALSE  actual=%lf\n", (double)__GET_VAR(data__->TESTBLOCK.NORTHSOUTHGREEN,));}
      {printf("2,0: TestBlock.EastWestRed = TRUE  actual=%lf\n", (double)__GET_VAR(data__->TESTBLOCK.EASTWESTRED,));}
      {printf("2,0: TestBlock.EastWestYellow = FALSE  actual=%lf\n", (double)__GET_VAR(data__->TESTBLOCK.EASTWESTYELLOW,));}
      {printf("2,0: TestBlock.EastWestGreen = TRUE  actual=%lf\n", (double)__GET_VAR(data__->TESTBLOCK.EASTWESTGREEN,));}
      {printf("2,0: TestBlock.PedestrianLight1 = FALSE  actual=%lf\n", (double)__GET_VAR(data__->TESTBLOCK.PEDESTRIANLIGHT1,));}
      {printf("2,0: TestBlock.PedestrianLight2 = TRUE  actual=%lf\n", (double)__GET_VAR(data__->TESTBLOCK.PEDESTRIANLIGHT2,));}
        IF NOT(TestBlock.NorthSouthRed = TRUE AND TestBlock.NorthSouthYellow = FALSE AND TestBlock.NorthSouthGreen = FALSE AND TestBlock.EastWestRed = TRUE AND TestBlock.EastWestYellow = FALSE AND TestBlock.EastWestGreen = TRUE AND TestBlock.PedestrianLight1 = FALSE AND TestBlock.PedestrianLight2 = TRUE) THEN Failed := TRUE; END_IF;
      END_IF;
      Finished:=TRUE;
  END_CASE;
END_FUNCTION_BLOCK

FUNCTION_BLOCK FB_TEST_3
  VAR_OUTPUT
    Finished : BOOL;
    Failed : BOOL;
  END_VAR
  VAR
    TestBlock : TRAFFIC_CTRL;
    TestState : INT;
    Timer : TON;
  END_VAR

  Timer(IN:=TRUE, PT:= T#0s); (* placeholder for later usage *)

  CASE testState OF
    0:
      IF (Timer.Q) THEN
        TestBlock(PedestrianButton1 := TRUE, PedestrianButton2 := TRUE);
        TestState:=TestState+1;
      END_IF;
      Timer(IN:=TRUE, PT:=T#0s);
    1:
      IF (Timer.Q) THEN
      {printf("3,0: TestBlock.NorthSouthRed = TRUE  actual=%lf\n", (double)__GET_VAR(data__->TESTBLOCK.NORTHSOUTHRED,));}
      {printf("3,0: TestBlock.NorthSouthYellow = FALSE  actual=%lf\n", (double)__GET_VAR(data__->TESTBLOCK.NORTHSOUTHYELLOW,));}
      {printf("3,0: TestBlock.NorthSouthGreen = FALSE  actual=%lf\n", (double)__GET_VAR(data__->TESTBLOCK.NORTHSOUTHGREEN,));}
      {printf("3,0: TestBlock.EastWestRed = TRUE  actual=%lf\n", (double)__GET_VAR(data__->TESTBLOCK.EASTWESTRED,));}
      {printf("3,0: TestBlock.EastWestYellow = TRUE  actual=%lf\n", (double)__GET_VAR(data__->TESTBLOCK.EASTWESTYELLOW,));}
      {printf("3,0: TestBlock.EastWestGreen = FALSE  actual=%lf\n", (double)__GET_VAR(data__->TESTBLOCK.EASTWESTGREEN,));}
      {printf("3,0: TestBlock.PedestrianLight1 = TRUE  actual=%lf\n", (double)__GET_VAR(data__->TESTBLOCK.PEDESTRIANLIGHT1,));}
      {printf("3,0: TestBlock.PedestrianLight2 = TRUE  actual=%lf\n", (double)__GET_VAR(data__->TESTBLOCK.PEDESTRIANLIGHT2,));}
        IF NOT(TestBlock.NorthSouthRed = TRUE AND TestBlock.NorthSouthYellow = FALSE AND TestBlock.NorthSouthGreen = FALSE AND TestBlock.EastWestRed = TRUE AND TestBlock.EastWestYellow = TRUE AND TestBlock.EastWestGreen = FALSE AND TestBlock.PedestrianLight1 = TRUE AND TestBlock.PedestrianLight2 = TRUE) THEN Failed := TRUE; END_IF;
      END_IF;
      Finished:=TRUE;
  END_CASE;
END_FUNCTION_BLOCK

PROGRAM TestRunnerProgram
VAR
  testResult AT %QX0.0 : BOOL := FALSE;
END_VAR
VAR
  totalTests AT %QW0 : INT := 0;
  passedTests AT %QW1 : INT := 0;
END_VAR
VAR
  i: INT := 0;
  testOutcomeArray : ARRAY [0..3] OF BOOL;
  Test_0: FB_TEST_0;
  Test_1: FB_TEST_1;
  Test_2: FB_TEST_2;
  Test_3: FB_TEST_3;
END_VAR

  IF NOT Test_0.Finished AND NOT Test_0.FAILED THEN totalTests := totalTests + 1; Test_0(); END_IF;
  IF Test_0.Finished THEN testOutcomeArray[0] := TRUE; END_IF;
  IF NOT Test_1.Finished AND NOT Test_1.FAILED THEN totalTests := totalTests + 1; Test_1(); END_IF;
  IF Test_1.Finished THEN testOutcomeArray[1] := TRUE; END_IF;
  IF NOT Test_2.Finished AND NOT Test_2.FAILED THEN totalTests := totalTests + 1; Test_2(); END_IF;
  IF Test_2.Finished THEN testOutcomeArray[2] := TRUE; END_IF;
  IF NOT Test_3.Finished AND NOT Test_3.FAILED THEN totalTests := totalTests + 1; Test_3(); END_IF;
  IF Test_3.Finished THEN testOutcomeArray[3] := TRUE; END_IF;

  passedTests := 0;
  FOR i:=0 TO 3 DO
    IF testOutcomeArray[i]=TRUE THEN passedTests := passedTests+1; END_IF;
  END_FOR;
END_PROGRAM
